FUNCTION_BLOCK PUMP_PROTECTION (* Migrated from IEC 61131-3 ST *)
  (* Standard: 61499-2 *)
  (* Version 1.0, 2026-11-06, st2fb *)
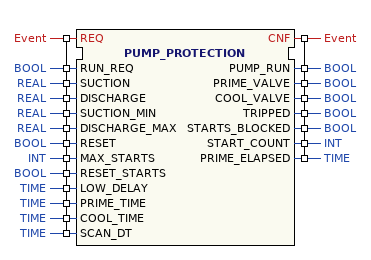
  EVENT_INPUT
    REQ WITH RUN_REQ, SUCTION, DISCHARGE, SUCTION_MIN, DISCHARGE_MAX, RESET, MAX_STARTS, RESET_STARTS, LOW_DELAY, PRIME_TIME, COOL_TIME, SCAN_DT;
  END_EVENT
  EVENT_OUTPUT
    CNF WITH PUMP_RUN, PRIME_VALVE, COOL_VALVE, TRIPPED, STARTS_BLOCKED, START_COUNT, PRIME_ELAPSED;
  END_EVENT
  VAR_INPUT
    RUN_REQ : BOOL;
    SUCTION : REAL;
    DISCHARGE : REAL;
    SUCTION_MIN : REAL;
    DISCHARGE_MAX : REAL;
    RESET : BOOL;
    MAX_STARTS : INT;
    RESET_STARTS : BOOL;
    LOW_DELAY : TIME;
    PRIME_TIME : TIME;
    COOL_TIME : TIME;
    SCAN_DT : TIME;
  END_VAR
  VAR_OUTPUT
    PUMP_RUN : BOOL;
    PRIME_VALVE : BOOL;
    COOL_VALVE : BOOL;
    TRIPPED : BOOL;
    STARTS_BLOCKED : BOOL;
    START_COUNT : INT;
    PRIME_ELAPSED : TIME;
  END_VAR
  VAR
    ST2FB_NOW : TIME := T#0s;
    RESTART_OK : BOOL;
    LOW_TIMER_IN : BOOL;
    LOW_TIMER_PT : TIME;
    LOW_TIMER_Q : BOOL;
    LOW_TIMER_ET : TIME;
    LOW_TIMER_STATE : INT;
    LOW_TIMER_PREV_IN : BOOL;
    LOW_TIMER_START_TIME : TIME;
    TRIP_LATCH_S : BOOL;
    TRIP_LATCH_R1 : BOOL;
    TRIP_LATCH_Q1 : BOOL;
    PRIME_PULSE_IN : BOOL;
    PRIME_PULSE_PT : TIME;
    PRIME_PULSE_Q : BOOL;
    PRIME_PULSE_ET : TIME;
    PRIME_PULSE_STATE : INT;
    PRIME_PULSE_PREV_IN : BOOL;
    PRIME_PULSE_START_TIME : TIME;
    COOL_DOWN_IN : BOOL;
    COOL_DOWN_PT : TIME;
    COOL_DOWN_Q : BOOL;
    COOL_DOWN_ET : TIME;
    COOL_DOWN_STATE : INT;
    COOL_DOWN_PREV_IN : BOOL;
    COOL_DOWN_START_TIME : TIME;
    START_COUNTER_CU : BOOL;
    START_COUNTER_R : BOOL;
    START_COUNTER_PV : INT;
    START_COUNTER_Q : BOOL;
    START_COUNTER_CV : INT;
    START_COUNTER_CU_T_Q : BOOL;
    START_COUNTER_CU_T_M : BOOL;
  END_VAR
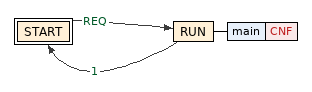
  EC_STATES
    START;
    RUN : main -> CNF;
  END_STATES
  EC_TRANSITIONS
    START TO RUN := REQ;
    RUN TO START := 1;
  END_TRANSITIONS
  ALGORITHM main IN ST:
ST2FB_NOW := ST2FB_NOW + SCAN_DT;

(* LOW_TIMER : TON *)
LOW_TIMER_IN := PUMP_RUN AND (SUCTION < SUCTION_MIN);
LOW_TIMER_PT := LOW_DELAY;
IF (LOW_TIMER_STATE = 0) AND NOT LOW_TIMER_PREV_IN AND LOW_TIMER_IN THEN
  LOW_TIMER_STATE := 1;
  LOW_TIMER_Q := FALSE;
  LOW_TIMER_START_TIME := ST2FB_NOW;
ELSE
  IF NOT LOW_TIMER_IN THEN
    LOW_TIMER_ET := T#0s;
    LOW_TIMER_Q := FALSE;
    LOW_TIMER_STATE := 0;
  ELSIF LOW_TIMER_STATE = 1 THEN
    IF LOW_TIMER_START_TIME + LOW_TIMER_PT <= ST2FB_NOW THEN
      LOW_TIMER_STATE := 2;
      LOW_TIMER_Q := TRUE;
      LOW_TIMER_ET := LOW_TIMER_PT;
    ELSE
      LOW_TIMER_ET := ST2FB_NOW - LOW_TIMER_START_TIME;
    END_IF;
  END_IF;
END_IF;
LOW_TIMER_PREV_IN := LOW_TIMER_IN;

(* TRIP_LATCH : RS *)
TRIP_LATCH_S := LOW_TIMER_Q OR (DISCHARGE > DISCHARGE_MAX);
TRIP_LATCH_R1 := RESET;
TRIP_LATCH_Q1 := NOT TRIP_LATCH_R1 AND (TRIP_LATCH_S OR TRIP_LATCH_Q1);
TRIPPED := TRIP_LATCH_Q1;
STARTS_BLOCKED := START_COUNTER_Q;
RESTART_OK := PUMP_RUN OR (NOT COOL_DOWN_Q AND NOT STARTS_BLOCKED);
PUMP_RUN := RUN_REQ AND NOT TRIPPED AND RESTART_OK;

(* START_COUNTER : CTU *)
START_COUNTER_CU := PUMP_RUN;
START_COUNTER_R := RESET_STARTS;
START_COUNTER_PV := MAX_STARTS;
START_COUNTER_CU_T_Q := START_COUNTER_CU AND NOT START_COUNTER_CU_T_M;
START_COUNTER_CU_T_M := START_COUNTER_CU;
IF START_COUNTER_R THEN
  START_COUNTER_CV := 0;
ELSIF START_COUNTER_CU_T_Q AND (START_COUNTER_CV < START_COUNTER_PV) THEN
  START_COUNTER_CV := START_COUNTER_CV + 1;
END_IF;
START_COUNTER_Q := START_COUNTER_CV >= START_COUNTER_PV;
START_COUNT := START_COUNTER_CV;

(* PRIME_PULSE : TP *)
PRIME_PULSE_IN := PUMP_RUN;
PRIME_PULSE_PT := PRIME_TIME;
IF (PRIME_PULSE_STATE = 0) AND NOT PRIME_PULSE_PREV_IN AND PRIME_PULSE_IN THEN
  PRIME_PULSE_STATE := 1;
  PRIME_PULSE_Q := TRUE;
  PRIME_PULSE_START_TIME := ST2FB_NOW;
ELSIF PRIME_PULSE_STATE = 1 THEN
  IF PRIME_PULSE_START_TIME + PRIME_PULSE_PT <= ST2FB_NOW THEN
    PRIME_PULSE_STATE := 2;
    PRIME_PULSE_Q := FALSE;
    PRIME_PULSE_ET := PRIME_PULSE_PT;
  ELSE
    PRIME_PULSE_ET := ST2FB_NOW - PRIME_PULSE_START_TIME;
  END_IF;
END_IF;
IF (PRIME_PULSE_STATE = 2) AND NOT PRIME_PULSE_IN THEN
  PRIME_PULSE_ET := T#0s;
  PRIME_PULSE_STATE := 0;
END_IF;
PRIME_PULSE_PREV_IN := PRIME_PULSE_IN;
PRIME_VALVE := PRIME_PULSE_Q;
PRIME_ELAPSED := PRIME_PULSE_ET;

(* COOL_DOWN : TOF *)
COOL_DOWN_IN := PUMP_RUN;
COOL_DOWN_PT := COOL_TIME;
IF (COOL_DOWN_STATE = 0) AND COOL_DOWN_PREV_IN AND NOT COOL_DOWN_IN THEN
  COOL_DOWN_STATE := 1;
  COOL_DOWN_START_TIME := ST2FB_NOW;
ELSE
  IF COOL_DOWN_IN THEN
    COOL_DOWN_ET := T#0s;
    COOL_DOWN_STATE := 0;
  ELSIF COOL_DOWN_STATE = 1 THEN
    IF COOL_DOWN_START_TIME + COOL_DOWN_PT <= ST2FB_NOW THEN
      COOL_DOWN_STATE := 2;
      COOL_DOWN_ET := COOL_DOWN_PT;
    ELSE
      COOL_DOWN_ET := ST2FB_NOW - COOL_DOWN_START_TIME;
    END_IF;
  END_IF;
END_IF;
COOL_DOWN_Q := COOL_DOWN_IN OR (COOL_DOWN_STATE = 1);
COOL_DOWN_PREV_IN := COOL_DOWN_IN;
COOL_VALVE := COOL_DOWN_Q;
  END_ALGORITHM
END_FUNCTION_BLOCK
